Fanuc KAREL source: KT00209.KL

PROGRAM KT00209
%NOLOCKGROUP
VAR
  Y1: ARRAY[2] OF BYTE
  B2: BOOLEAN
  OUT: BOOLEAN
BEGIN
  Y1[1] = 2
    B2 = FALSE
  OUT = Y1[1] AND B2
END KT00209
